Yaskawa INFORM job: HAND_CLOSE.JBI

/JOB
//NAME HAND_CLOSE
//POS
///NPOS 0,0,0,0,0,0
//INST
///DATE 2026/10/09 19:37
///COMM GRIPPER CLOSE
///ATTR SC,RW
NOP
DOUT OT#(2) OFF
DOUT OT#(1) ON
WAIT IN#(1)=ON T=3.00
TIMER T=0.20
END
